(*
SPDX-FileCopyrightText: c 2026 Oleksandr Tiutyk <trofimich@gmail.com>
SPDX-License-Identifier: MIT
License: https://opensource.org/license/mit
*)

(*!
<summary>Checks prefix/value/suffix order and callback counts.</summary>
<description>
Owns persistent native serializer state and any payload buffers used by this case.
Run from one task at a stable address. The caller provides task-boundary exception cleanup.
</description>
*)

{attribute 'no_assign'}
{attribute 'no_explicit_call' := 'do not call this function block directly'}
FUNCTION_BLOCK AutomaticJsonWrappedCallbacksTest EXTENDS TOF_Testing.SingleCycleTest
VAR_STAT
	{attribute 'hide'}
	_ClassName : STRING := __POUNAME();
END_VAR
VAR
	_Serializer : TOF_JSON.AutomaticJsonSerializer;
	_Extender : JsonExtenderProbe;
	_Source : JSON_TEST_VALUE;
	_Json : TOF_Core.JSON_DOCUMENT;
END_VAR

(*!
<summary>Checks prefix/value/suffix order and callback counts.</summary>
*)
METHOD PROTECTED ExecuteTest
VAR
	success : BOOL;
	jsonSize : UDINT;
	expectedJson : STRING(40) := '[{"Number":42,"Ready":true}]';
END_VAR
_Source.Number := 42;
_Source.Ready := TRUE;

_Json := '';

_Extender.Reset();

success := _Serializer.TrySerialize(
	sourceStructure := _Source,
	extender := _Extender,
	targetJson := _Json,
	jsonSize => jsonSize
);
Assert.ThatBool(
	actual := success,
	message := "Balanced callbacks must produce a document"
).IsTrue();
Assert.That(
	actual := _Json,
	message := "Callbacks must surround exactly one structure value"
).ToBe(expected := expectedJson);
Assert.ThatUDInt(
	actual := _Extender.StartCount,
	message := "Start must run once"
).ToBe(expected := 1);
Assert.ThatUDInt(
	actual := _Extender.FinishCount,
	message := "Finish must run once"
).ToBe(expected := 1);
END_METHOD

(*!
<summary>Restores the fixture before the runner publishes the result.</summary>
<description>
Also runs after an unexpected exception interrupts the case.
</description>
*)
METHOD PROTECTED AfterTest
_Extender.Reset();
END_METHOD

//! <summary>Borrows the concrete class name. Callers must not modify it.</summary>
{attribute 'monitoring' := 'call'}
PROPERTY ClassName : REFERENCE TO STRING
GET
ClassName REF= _ClassName;
END_GET
END_PROPERTY

//! <summary>Borrows the compiler-initialized namespace name. Callers must not modify it.</summary>
{attribute 'monitoring' := 'call'}
PROPERTY NamespaceName : REFERENCE TO STRING
GET
NamespaceName REF= CurrentNamespace.Name;
END_GET
END_PROPERTY

//! <summary>Reports the concrete instance size in bytes.</summary>
{attribute 'monitoring' := 'call'}
PROPERTY SelfSize : ULINT
GET
SelfSize := XSIZEOF(THIS^);
END_GET
END_PROPERTY

END_FUNCTION_BLOCK

(* stored: Version 1.1.0.1
   POU AutomaticJsonWrappedCallbacksTest: Id {c677a228-f281-43da-a5f4-5b5c488b19d8}, SpecialFunc None
   Method ExecuteTest: Id {4406ba9c-761e-4566-aa70-94f24142f07c}
   Method AfterTest: Id {50c15499-3d63-4910-81be-1add4158f330}
   Property ClassName: Id {64a2328c-dfb6-465a-aa42-948b208c2cf8}
   Get Get: Id {12f0d956-a1f3-49b2-815f-5b048ec3aafd}
   Property NamespaceName: Id {cd5dacb1-ada8-435f-8c8c-3d9057ee00d0}
   Get Get: Id {0f0b4bd5-fd2b-461c-8224-f435f6518952}
   Property SelfSize: Id {75580b33-03ec-449c-bc8e-b91745a8cb8e}
   Get Get: Id {ed6c6f29-8221-4d17-bc52-9c19e7e2006b} *)
